        pointRx pPointRx[2] = {x=594.549819, y=30.770866, z=171.45682, rx=-40.410864, ry=94.502866, rz=40.920287, shoulder=lefty, elbow=epositive, wrist=wnegative}
        string sID
      [28]
        bool bMarked
        jointRx jJointRx = {j1=-1.639134, j2=22.193742, j3=116.03978, j4=1.817031, j5=-44.819098, j6=-0.790246}
        pointRx pInter
        paraItem pParaItem
          [0]
            bool bSafePoint
            ifItem iIfItem
              [0]
                bool bANDOR[2]
                num nSigIndex[3]
                num nSigType[3]
                num nValue[3]
            mdesc mMdesc = {accel=25, vel=50, leave=1}
            num nActionIndex = 8
            num nDelay = 1.2
            num nMoveType = 7
            num nPercentage
            num nSigValue = 1
        pointRx pPointRx[2] = {x=594.549757, y=30.770873, z=70.540177, rx=-40.399083, ry=94.503271, rz=40.908669, shoulder=lefty, elbow=epositive, wrist=wnegative}
        string sID
      [29]
        bool bMarked
        jointRx jJointRx = {j1=-1.639045, j2=12.402747, j3=111.595585, j4=2.517874, j5=-30.594648, j6=-1.669011}
        pointRx pInter
        paraItem pParaItem
          [0]
            bool bSafePoint
            ifItem iIfItem
              [0]
                bool bANDOR[2]
                num nSigIndex[3]
                num nSigType[3]
                num nValue[3]
            mdesc mMdesc
            num nActionIndex = 10
            num nDelay = 5
            num nMoveType = 4
            num nPercentage
            num nSigValue
        pointRx pPointRx[2] = {x=594.549819, y=30.770866, z=171.45682, rx=-40.410864, ry=94.502866, rz=40.920287, shoulder=lefty, elbow=epositive, wrist=wnegative}
        string sID
      [30]
        bool bMarked
        jointRx jJointRx = {j1=-1.639045, j2=12.402747, j3=111.595585, j4=2.517874, j5=-30.594648, j6=-1.669011}
        pointRx pInter
        paraItem pParaItem
          [0]
            bool bSafePoint
            ifItem iIfItem
              [0]
                bool bANDOR[2]
                num nSigIndex[3]
                num nSigType[3]
                num nValue[3]
            mdesc mMdesc
            num nActionIndex = 10
            num nDelay = 0.5
            num nMoveType = 7
            num nPercentage
            num nSigValue
        pointRx pPointRx[2] = {x=594.549819, y=30.770866, z=171.45682, rx=-40.410864, ry=94.502866, rz=40.920287, shoulder=lefty, elbow=epositive, wrist=wnegative}
        string sID
      [31]
        bool bMarked
        jointRx jJointRx = {j1=-1.639045, j2=12.402747, j3=111.595585, j4=2.517874, j5=-30.594648, j6=-1.669011}
        pointRx pInter
        paraItem pParaItem
          [0]
            bool bSafePoint
            ifItem iIfItem
              [0]
                bool bANDOR[2]
                num nSigIndex[3]
                num nSigType[3]
                num nValue[3]
            mdesc mMdesc
            num nActionIndex = 9
            num nDelay = 5
            num nMoveType = 3
            num nPercentage
            num nSigValue = 1
        pointRx pPointRx[2] = {x=594.549819, y=30.770866, z=171.45682, rx=-40.410864, ry=94.502866, rz=40.920287, shoulder=lefty, elbow=epositive, wrist=wnegative}
        string sID
      [32]
        bool bMarked
        jointRx jJointRx = {j1=-7.226415, j2=23.592658, j3=117.966616, j4=-6.814076, j5=-74.706283, j6=4.672196}
        pointRx pInter
        paraItem pParaItem
          [0]
            bool bSafePoint
            ifItem iIfItem
              [0]
                bool bANDOR[2]
                num nSigIndex[3]
                num nSigType[3]
                num nValue[3]
            mdesc mMdesc
            num nActionIndex = 9
            num nDelay = 5
            num nMoveType
            num nPercentage
            num nSigValue = 1
        pointRx pPointRx[2] = {x=578.895133, y=-11.466034, z=95.479539, rx=0.214531, ry=67.116514, rz=-0.152975, shoulder=lefty, elbow=epositive, wrist=wnegative}
        string sID
      [33]
        bool bMarked
        jointRx jJointRx = {j1=-2.687248, j2=16.117165, j3=122.304638, j4=-0.487867, j5=-66.528565, j6=1.978834}
        pointRx pInter
        paraItem pParaItem
          [0]
            bool bSafePoint
            ifItem iIfItem
              [0]
                bool bANDOR[2]
                num nSigIndex[3]
                num nSigType[3]
                num nValue[3]
            mdesc mMdesc
            num nActionIndex = 1
            num nDelay = 5
            num nMoveType = 6
            num nPercentage
            num nSigValue = 1
        pointRx pPointRx[2] = {x=546.855577, y=25.169852, z=121.450925, rx=6.745985, ry=71.76392, rz=-5.460967, shoulder=lefty, elbow=epositive, wrist=wnegative}
        string sID
      [34]
        bool bMarked
        jointRx jJointRx = {j1=-2.687248, j2=16.117165, j3=122.304638, j4=-0.487867, j5=-66.528565, j6=1.978834}
        pointRx pInter
        paraItem pParaItem
          [0]
            bool bSafePoint
            ifItem iIfItem
              [0]
                bool bANDOR[2]
                num nSigIndex[3]
                num nSigType[3]
                num nValue[3]
            mdesc mMdesc
            num nActionIndex = 1
            num nDelay = 5
            num nMoveType = 5
            num nPercentage
            num nSigValue = 1
        pointRx pPointRx[2] = {x=546.855577, y=25.169852, z=121.450925, rx=6.745985, ry=71.76392, rz=-5.460967, shoulder=lefty, elbow=epositive, wrist=wnegative}
        string sID
      [35]
        bool bMarked
        jointRx jJointRx = {j1=-1.639045, j2=12.402747, j3=111.595585, j4=2.517874, j5=-30.594648, j6=-1.669011}
        pointRx pInter
        paraItem pParaItem
          [0]
            bool bSafePoint
            ifItem iIfItem
              [0]
                bool bANDOR[2]
                num nSigIndex[3]
                num nSigType[3]
                num nValue[3]
            mdesc mMdesc
            num nActionIndex = 10
            num nDelay
            num nMoveType = 4
            num nPercentage
            num nSigValue = 1
        pointRx pPointRx[2] = {x=594.549819, y=30.770866, z=171.45682, rx=-40.410864, ry=94.502866, rz=40.920287, shoulder=lefty, elbow=epositive, wrist=wnegative}
        string sID
      [36]
        bool bMarked
        jointRx jJointRx = {j1=-1.639045, j2=12.402747, j3=111.595585, j4=2.517874, j5=-30.594648, j6=-1.669011}
        pointRx pInter
        paraItem pParaItem
          [0]
            bool bSafePoint
            ifItem iIfItem
              [0]
                bool bANDOR[2]
                num nSigIndex[3]
                num nSigType[3]
                num nValue[3]
            mdesc mMdesc
            num nActionIndex = 8
            num nDelay
            num nMoveType = 3
            num nPercentage
            num nSigValue = 1
        pointRx pPointRx[2] = {x=594.549819, y=30.770866, z=171.45682, rx=-40.410864, ry=94.502866, rz=40.920287, shoulder=lefty, elbow=epositive, wrist=wnegative}
        string sID
      [37]
        bool bMarked
        jointRx jJointRx = {j1=-1.639134, j2=22.193742, j3=116.03978, j4=1.817031, j5=-44.819098, j6=-0.790246}
        pointRx pInter
        paraItem pParaItem
          [0]
            bool bSafePoint
            ifItem iIfItem
              [0]
                bool bANDOR[2]
                num nSigIndex[3]
                num nSigType[3]
                num nValue[3]
            mdesc mMdesc = {accel=25, vel=50, leave=1}
            num nActionIndex = 8
            num nDelay = 1.2
            num nMoveType = 7
            num nPercentage
            num nSigValue = 1
        pointRx pPointRx[2] = {x=594.549757, y=30.770873, z=70.540177, rx=-40.399083, ry=94.503271, rz=40.908669, shoulder=lefty, elbow=epositive, wrist=wnegative}
        string sID
      [38]
        bool bMarked
        jointRx jJointRx = {j1=-1.639045, j2=12.402747, j3=111.595585, j4=2.517874, j5=-30.594648, j6=-1.669011}
        pointRx pInter
        paraItem pParaItem
          [0]
            bool bSafePoint
            ifItem iIfItem
              [0]
                bool bANDOR[2]
                num nSigIndex[3]
                num nSigType[3]
                num nValue[3]
            mdesc mMdesc
            num nActionIndex = 10
            num nDelay = 5
            num nMoveType = 4
            num nPercentage
            num nSigValue
        pointRx pPointRx[2] = {x=594.549819, y=30.770866, z=171.45682, rx=-40.410864, ry=94.502866, rz=40.920287, shoulder=lefty, elbow=epositive, wrist=wnegative}
        string sID
      [39]
        bool bMarked
        jointRx jJointRx = {j1=-1.639045, j2=12.402747, j3=111.595585, j4=2.517874, j5=-30.594648, j6=-1.669011}
        pointRx pInter
        paraItem pParaItem
          [0]
            bool bSafePoint
            ifItem iIfItem
              [0]
                bool bANDOR[2]
                num nSigIndex[3]
                num nSigType[3]
                num nValue[3]
            mdesc mMdesc
            num nActionIndex = 10
            num nDelay = 0.5
            num nMoveType = 7
            num nPercentage
            num nSigValue
        pointRx pPointRx[2] = {x=594.549819, y=30.770866, z=171.45682, rx=-40.410864, ry=94.502866, rz=40.920287, shoulder=lefty, elbow=epositive, wrist=wnegative}
        string sID
      [40]
        bool bMarked
        jointRx jJointRx = {j1=-1.639045, j2=12.402747, j3=111.595585, j4=2.517874, j5=-30.594648, j6=-1.669011}
        pointRx pInter
        paraItem pParaItem
          [0]
            bool bSafePoint
            ifItem iIfItem
              [0]
                bool bANDOR[2]
                num nSigIndex[3]
                num nSigType[3]
                num nValue[3]
            mdesc mMdesc
            num nActionIndex = 9
            num nDelay = 5
            num nMoveType = 3
            num nPercentage
            num nSigValue = 1
        pointRx pPointRx[2] = {x=594.549819, y=30.770866, z=171.45682, rx=-40.410864, ry=94.502866, rz=40.920287, shoulder=lefty, elbow=epositive, wrist=wnegative}
        string sID
      [41]
        bool bMarked
        jointRx jJointRx = {j1=-5.695731, j2=1.0651158, j3=140.857781, j4=-5.0995594, j5=-70.16665, j6=4.945113}
        pointRx pInter
        paraItem pParaItem
          [0]
            bool bSafePoint
            ifItem iIfItem
              [0]
                bool bANDOR[2]
                num nSigIndex[3]
                num nSigType[3]
                num nValue[3]
            mdesc mMdesc
            num nActionIndex = 9
            num nDelay = 5
            num nMoveType
            num nPercentage
            num nSigValue = 1
        pointRx pPointRx[2] = {x=418.431788, y=16.917425, z=121.450805, rx=1.98388, ry=71.88349, rz=-0.448462, shoulder=lefty, elbow=epositive, wrist=wnegative}
        string sID
      [42]
        bool bMarked
        jointRx jJointRx = {j1=-7.298028, j2=2.858926, j3=83.785178, j4=10.154119, j5=40.0244602, j6=-11.233253}
        pointRx pInter
        paraItem pParaItem
          [0]
            bool bSafePoint
            ifItem iIfItem
              [0]
                bool bANDOR[2]
                num nSigIndex[3]
                num nSigType[3]
                num nValue[3]
            mdesc mMdesc
            num nActionIndex = 9
            num nDelay = 5
            num nMoveType
            num nPercentage
            num nSigValue = 1
        pointRx pPointRx[2] = {x=578.748864, y=-12.280333, z=390.636728, rx=1.0385678, ry=125.960392, rz=0.0408503, shoulder=lefty, elbow=epositive, wrist=wpositive}
        string sID
      [43]
        bool bMarked
        jointRx jJointRx = {j1=-11.714441, j2=6.765338, j3=77.722005, j4=11.0036166, j5=46.0689495, j6=-14.380804}
        pointRx pInter
        paraItem pParaItem
          [0]
            bool bSafePoint
            ifItem iIfItem
              [0]
                bool bANDOR[2]
                num nSigIndex[3]
                num nSigType[3]
                num nValue[3]
            mdesc mMdesc
            num nActionIndex = 1
            num nDelay = 5
            num nMoveType = 6
            num nPercentage
            num nSigValue = 1
        pointRx pPointRx[2] = {x=599.417794, y=-59.189006, z=399.167028, rx=-1.744645, ry=129.591612, rz=2.151169, shoulder=lefty, elbow=epositive, wrist=wpositive}
        string sID
      [44]
        bool bMarked
        jointRx jJointRx = {j1=-11.714441, j2=6.765338, j3=77.722005, j4=11.0036166, j5=46.0689495, j6=-14.380804}
        pointRx pInter
        paraItem pParaItem
          [0]
            bool bSafePoint
            ifItem iIfItem
              [0]
                bool bANDOR[2]
                num nSigIndex[3]
                num nSigType[3]
                num nValue[3]
            mdesc mMdesc
            num nActionIndex = 1
            num nDelay = 5
            num nMoveType = 5
            num nPercentage
            num nSigValue = 1
        pointRx pPointRx[2] = {x=599.417794, y=-59.189006, z=399.167028, rx=-1.744645, ry=129.591612, rz=2.151169, shoulder=lefty, elbow=epositive, wrist=wpositive}
        string sID
      [45]
        bool bMarked
        jointRx jJointRx = {j1=-11.714441, j2=6.765338, j3=77.722005, j4=11.0036166, j5=46.0689495, j6=-14.380804}
        pointRx pInter
        paraItem pParaItem
          [0]
            bool bSafePoint
            ifItem iIfItem
              [0]
                bool bANDOR[2]
                num nSigIndex[3]
                num nSigType[3]
                num nValue[3]
            mdesc mMdesc
            num nActionIndex = 10
            num nDelay = 5
            num nMoveType = 4
            num nPercentage
            num nSigValue = 1
        pointRx pPointRx[2] = {x=599.417794, y=-59.189006, z=399.167028, rx=-1.744645, ry=129.591612, rz=2.151169, shoulder=lefty, elbow=epositive, wrist=wpositive}
        string sID
      [46]
        bool bMarked
        jointRx jJointRx = {j1=-11.714441, j2=6.765338, j3=77.722005, j4=11.0036166, j5=46.0689495, j6=-14.380804}
        pointRx pInter
        paraItem pParaItem
          [0]
            bool bSafePoint
            ifItem iIfItem
              [0]
                bool bANDOR[2]
                num nSigIndex[3]
                num nSigType[3]
                num nValue[3]
            mdesc mMdesc
            num nActionIndex = 8
            num nDelay = 5
            num nMoveType = 3
            num nPercentage
            num nSigValue = 1
        pointRx pPointRx[2] = {x=599.417794, y=-59.189006, z=399.167028, rx=-1.744645, ry=129.591612, rz=2.151169, shoulder=lefty, elbow=epositive, wrist=wpositive}
        string sID
      [47]
        bool bMarked
        jointRx jJointRx = {j1=-11.714441, j2=6.765338, j3=77.722005, j4=11.0036166, j5=46.0689495, j6=-14.380804}
        pointRx pInter
        paraItem pParaItem
          [0]
            bool bSafePoint
            ifItem iIfItem
              [0]
                bool bANDOR[2]
                num nSigIndex[3]
                num nSigType[3]
                num nValue[3]
            mdesc mMdesc
            num nActionIndex = 8
            num nDelay = 2
            num nMoveType = 7
            num nPercentage
            num nSigValue = 1
        pointRx pPointRx[2] = {x=599.417794, y=-59.189006, z=399.167028, rx=-1.744645, ry=129.591612, rz=2.151169, shoulder=lefty, elbow=epositive, wrist=wpositive}
        string sID
      [48]
        bool bMarked
        jointRx jJointRx = {j1=-11.714441, j2=6.765338, j3=77.722005, j4=11.0036166, j5=46.0689495, j6=-14.380804}
        pointRx pInter
        paraItem pParaItem
          [0]
            bool bSafePoint
            ifItem iIfItem
              [0]
                bool bANDOR[2]
                num nSigIndex[3]
                num nSigType[3]
                num nValue[3]
            mdesc mMdesc
            num nActionIndex = 10
            num nDelay = 1
            num nMoveType = 4
            num nPercentage
            num nSigValue
        pointRx pPointRx[2] = {x=599.417794, y=-59.189006, z=399.167028, rx=-1.744645, ry=129.591612, rz=2.151169, shoulder=lefty, elbow=epositive, wrist=wpositive}
        string sID
      [49]
        bool bMarked
        jointRx jJointRx = {j1=-11.714441, j2=6.765338, j3=77.722005, j4=11.0036166, j5=46.0689495, j6=-14.380804}
        pointRx pInter
        paraItem pParaItem
          [0]
            bool bSafePoint
            ifItem iIfItem
              [0]
                bool bANDOR[2]
                num nSigIndex[3]
                num nSigType[3]
                num nValue[3]
            mdesc mMdesc
            num nActionIndex = 10
            num nDelay = 0.5
            num nMoveType = 7
            num nPercentage
            num nSigValue
        pointRx pPointRx[2] = {x=599.417794, y=-59.189006, z=399.167028, rx=-1.744645, ry=129.591612, rz=2.151169, shoulder=lefty, elbow=epositive, wrist=wpositive}
        string sID
      [50]
        bool bMarked
        jointRx jJointRx = {j1=-11.714441, j2=6.765338, j3=77.722005, j4=11.0036166, j5=46.0689495, j6=-14.380804}
        pointRx pInter
        paraItem pParaItem
          [0]
            bool bSafePoint
            ifItem iIfItem
              [0]
                bool bANDOR[2]
                num nSigIndex[3]
                num nSigType[3]
                num nValue[3]
            mdesc mMdesc
            num nActionIndex = 9
            num nDelay = 1
            num nMoveType = 3
            num nPercentage
            num nSigValue = 1
        pointRx pPointRx[2] = {x=599.417794, y=-59.189006, z=399.167028, rx=-1.744645, ry=129.591612, rz=2.151169, shoulder=lefty, elbow=epositive, wrist=wpositive}
        string sID
      [51]
        bool bMarked
        jointRx jJointRx = {j1=-1.121423, j2=3.0557806, j3=83.578223, j4=2.394681, j5=39.358319, j6=-1.629384}
        pointRx pInter
        paraItem pParaItem
          [0]
            bool bSafePoint
            ifItem iIfItem
              [0]
                bool bANDOR[2]
                num nSigIndex[3]
                num nSigType[3]
                num nValue[3]
            mdesc mMdesc
            num nActionIndex = 9
            num nDelay = 5
            num nMoveType
            num nPercentage
            num nSigValue = 1
        pointRx pPointRx[2] = {x=578.748846, y=41.330803, z=390.636723, rx=1.0399619, ry=125.960028, rz=0.0394555, shoulder=lefty, elbow=epositive, wrist=wpositive}
        string sID
      [52]
        bool bMarked
        jointRx jJointRx = {j1=-2.687248, j2=16.117165, j3=122.304638, j4=-0.487867, j5=-66.528565, j6=1.978834}
        pointRx pInter
        paraItem pParaItem
          [0]
            bool bSafePoint
            ifItem iIfItem
              [0]
                bool bANDOR[2]
                num nSigIndex[3]
                num nSigType[3]
                num nValue[3]
            mdesc mMdesc
            num nActionIndex = 1
            num nDelay = 5
            num nMoveType = 6
            num nPercentage
            num nSigValue = 1
        pointRx pPointRx[2] = {x=546.855577, y=25.169852, z=121.450925, rx=6.745985, ry=71.76392, rz=-5.460967, shoulder=lefty, elbow=epositive, wrist=wnegative}
        string sID
      [53]
        bool bMarked
        jointRx jJointRx = {j1=-2.687248, j2=16.117165, j3=122.304638, j4=-0.487867, j5=-66.528565, j6=1.978834}
        pointRx pInter
        paraItem pParaItem
          [0]
            bool bSafePoint
            ifItem iIfItem
              [0]
                bool bANDOR[2]
                num nSigIndex[3]
                num nSigType[3]
                num nValue[3]
            mdesc mMdesc
            num nActionIndex = 1
            num nDelay = 5
            num nMoveType = 5
            num nPercentage
            num nSigValue = 1
        pointRx pPointRx[2] = {x=546.855577, y=25.169852, z=121.450925, rx=6.745985, ry=71.76392, rz=-5.460967, shoulder=lefty, elbow=epositive, wrist=wnegative}
        string sID
      [54]
        bool bMarked
        jointRx jJointRx = {j1=-1.639045, j2=12.402747, j3=111.595585, j4=2.517874, j5=-30.594648, j6=-1.669011}
        pointRx pInter
        paraItem pParaItem
          [0]
            bool bSafePoint
            ifItem iIfItem
              [0]
                bool bANDOR[2]
                num nSigIndex[3]
                num nSigType[3]
                num nValue[3]
            mdesc mMdesc
            num nActionIndex = 10
            num nDelay
            num nMoveType = 4
            num nPercentage
            num nSigValue = 1
        pointRx pPointRx[2] = {x=594.549819, y=30.770866, z=171.45682, rx=-40.410864, ry=94.502866, rz=40.920287, shoulder=lefty, elbow=epositive, wrist=wnegative}
        string sID
      [55]
        bool bMarked
        jointRx jJointRx = {j1=-1.639045, j2=12.402747, j3=111.595585, j4=2.517874, j5=-30.594648, j6=-1.669011}
        pointRx pInter
        paraItem pParaItem
          [0]
            bool bSafePoint
            ifItem iIfItem
              [0]
                bool bANDOR[2]
                num nSigIndex[3]
                num nSigType[3]
                num nValue[3]
            mdesc mMdesc
            num nActionIndex = 8
            num nDelay
            num nMoveType = 3
            num nPercentage
            num nSigValue = 1
        pointRx pPointRx[2] = {x=594.549819, y=30.770866, z=171.45682, rx=-40.410864, ry=94.502866, rz=40.920287, shoulder=lefty, elbow=epositive, wrist=wnegative}
        string sID
      [56]
        bool bMarked
        jointRx jJointRx = {j1=-1.639134, j2=22.193742, j3=116.03978, j4=1.817031, j5=-44.819098, j6=-0.790246}
        pointRx pInter
        paraItem pParaItem
          [0]
            bool bSafePoint
            ifItem iIfItem
              [0]
                bool bANDOR[2]
                num nSigIndex[3]
                num nSigType[3]
                num nValue[3]
            mdesc mMdesc = {accel=25, vel=50, leave=1}
            num nActionIndex = 8
            num nDelay = 2
            num nMoveType = 7
            num nPercentage
            num nSigValue = 1
        pointRx pPointRx[2] = {x=594.549757, y=30.770873, z=70.540177, rx=-40.399083, ry=94.503271, rz=40.908669, shoulder=lefty, elbow=epositive, wrist=wnegative}
        string sID
      [57]
        bool bMarked
        jointRx jJointRx = {j1=-1.639045, j2=12.402747, j3=111.595585, j4=2.517874, j5=-30.594648, j6=-1.669011}
        pointRx pInter
        paraItem pParaItem
          [0]
            bool bSafePoint
            ifItem iIfItem
              [0]
                bool bANDOR[2]
                num nSigIndex[3]
                num nSigType[3]
                num nValue[3]
            mdesc mMdesc
            num nActionIndex = 10
            num nDelay = 5
            num nMoveType = 4
            num nPercentage
            num nSigValue
        pointRx pPointRx[2] = {x=594.549819, y=30.770866, z=171.45682, rx=-40.410864, ry=94.502866, rz=40.920287, shoulder=lefty, elbow=epositive, wrist=wnegative}
        string sID
      [58]
        bool bMarked
        jointRx jJointRx = {j1=-1.639045, j2=12.402747, j3=111.595585, j4=2.517874, j5=-30.594648, j6=-1.669011}
        pointRx pInter
        paraItem pParaItem
          [0]
            bool bSafePoint
            ifItem iIfItem
              [0]
                bool bANDOR[2]
                num nSigIndex[3]
                num nSigType[3]
                num nValue[3]
            mdesc mMdesc
            num nActionIndex = 10
            num nDelay = 0.5
            num nMoveType = 7
            num nPercentage
            num nSigValue
        pointRx pPointRx[2] = {x=594.549819, y=30.770866, z=171.45682, rx=-40.410864, ry=94.502866, rz=40.920287, shoulder=lefty, elbow=epositive, wrist=wnegative}
        string sID
      [59]
        bool bMarked
        jointRx jJointRx = {j1=-1.639045, j2=12.402747, j3=111.595585, j4=2.517874, j5=-30.594648, j6=-1.669011}
        pointRx pInter
        paraItem pParaItem
          [0]
            bool bSafePoint
            ifItem iIfItem
              [0]
                bool bANDOR[2]
                num nSigIndex[3]
                num nSigType[3]
                num nValue[3]
            mdesc mMdesc
            num nActionIndex = 9
            num nDelay = 5
            num nMoveType = 3
            num nPercentage
            num nSigValue = 1
        pointRx pPointRx[2] = {x=594.549819, y=30.770866, z=171.45682, rx=-40.410864, ry=94.502866, rz=40.920287, shoulder=lefty, elbow=epositive, wrist=wnegative}
        string sID
      [60]
        bool bMarked
        jointRx jJointRx = {j1=-3.420163, j2=22.945404, j3=44.641192, j4=2.309583, j5=82.959552, j6=-2.373603}
        pointRx pInter
        paraItem pParaItem
          [0]
            bool bSafePoint
            ifItem iIfItem
              [0]
                bool bANDOR[2]
                num nSigIndex[3]
                num nSigType[3]
                num nValue[3]
            mdesc mMdesc
            num nActionIndex = 9
            num nDelay = 5
            num nMoveType
            num nPercentage
            num nSigValue = 1
        pointRx pPointRx[2] = {x=659.773544, y=14.665083, z=466.418783, rx=0.698518, ry=150.466936, rz=0.542991, shoulder=lefty, elbow=epositive, wrist=wpositive}
        string sID
      [61]
        bool bMarked
        jointRx jJointRx = {j1=-2.687248, j2=16.117165, j3=122.304638, j4=-0.487867, j5=-66.528565, j6=1.978834}
        pointRx pInter
        paraItem pParaItem
          [0]
            bool bSafePoint
            ifItem iIfItem
              [0]
                bool bANDOR[2]
                num nSigIndex[3]
                num nSigType[3]
                num nValue[3]
            mdesc mMdesc
            num nActionIndex = 1
            num nDelay = 5
            num nMoveType = 6
            num nPercentage
            num nSigValue = 1
        pointRx pPointRx[2] = {x=546.855577, y=25.169852, z=121.450925, rx=6.745985, ry=71.76392, rz=-5.460967, shoulder=lefty, elbow=epositive, wrist=wnegative}
        string sID
      [62]
        bool bMarked
        jointRx jJointRx = {j1=-2.687248, j2=16.117165, j3=122.304638, j4=-0.487867, j5=-66.528565, j6=1.978834}
        pointRx pInter
        paraItem pParaItem
          [0]
            bool bSafePoint
            ifItem iIfItem
              [0]
                bool bANDOR[2]
                num nSigIndex[3]
                num nSigType[3]
                num nValue[3]
            mdesc mMdesc
            num nActionIndex = 1
            num nDelay = 5
            num nMoveType = 5
            num nPercentage
            num nSigValue = 1
        pointRx pPointRx[2] = {x=546.855577, y=25.169852, z=121.450925, rx=6.745985, ry=71.76392, rz=-5.460967, shoulder=lefty, elbow=epositive, wrist=wnegative}
        string sID
      [63]
        bool bMarked
        jointRx jJointRx = {j1=-1.639045, j2=12.402747, j3=111.595585, j4=2.517874, j5=-30.594648, j6=-1.669011}
        pointRx pInter
        paraItem pParaItem
          [0]
            bool bSafePoint
            ifItem iIfItem
              [0]
                bool bANDOR[2]
                num nSigIndex[3]
                num nSigType[3]
                num nValue[3]
            mdesc mMdesc
            num nActionIndex = 10
            num nDelay
            num nMoveType = 4
            num nPercentage
            num nSigValue = 1
        pointRx pPointRx[2] = {x=594.549819, y=30.770866, z=171.45682, rx=-40.410864, ry=94.502866, rz=40.920287, shoulder=lefty, elbow=epositive, wrist=wnegative}
        string sID
      [64]
        bool bMarked
        jointRx jJointRx = {j1=-1.639045, j2=12.402747, j3=111.595585, j4=2.517874, j5=-30.594648, j6=-1.669011}
        pointRx pInter
        paraItem pParaItem
          [0]
            bool bSafePoint
            ifItem iIfItem
              [0]
                bool bANDOR[2]
                num nSigIndex[3]
                num nSigType[3]
                num nValue[3]
            mdesc mMdesc
            num nActionIndex = 8
            num nDelay
            num nMoveType = 3
            num nPercentage
            num nSigValue = 1
        pointRx pPointRx[2] = {x=594.549819, y=30.770866, z=171.45682, rx=-40.410864, ry=94.502866, rz=40.920287, shoulder=lefty, elbow=epositive, wrist=wnegative}
        string sID
      [65]
        bool bMarked
        jointRx jJointRx = {j1=-1.639134, j2=22.193742, j3=116.03978, j4=1.817031, j5=-44.819098, j6=-0.790246}
        pointRx pInter
        paraItem pParaItem
          [0]
            bool bSafePoint
            ifItem iIfItem
              [0]
                bool bANDOR[2]
                num nSigIndex[3]
                num nSigType[3]
                num nValue[3]
            mdesc mMdesc = {accel=25, vel=50, leave=1}
            num nActionIndex = 8
            num nDelay = 1.2
            num nMoveType = 7
            num nPercentage
            num nSigValue = 1
        pointRx pPointRx[2] = {x=594.549757, y=30.770873, z=70.540177, rx=-40.399083, ry=94.503271, rz=40.908669, shoulder=lefty, elbow=epositive, wrist=wnegative}
        string sID
      [66]
        bool bMarked
        jointRx jJointRx = {j1=-1.639045, j2=12.402747, j3=111.595585, j4=2.517874, j5=-30.594648, j6=-1.669011}
        pointRx pInter
        paraItem pParaItem
          [0]
            bool bSafePoint
            ifItem iIfItem
              [0]
                bool bANDOR[2]
                num nSigIndex[3]
                num nSigType[3]
                num nValue[3]
            mdesc mMdesc
            num nActionIndex = 10
            num nDelay = 5
            num nMoveType = 4
            num nPercentage
            num nSigValue
        pointRx pPointRx[2] = {x=594.549819, y=30.770866, z=171.45682, rx=-40.410864, ry=94.502866, rz=40.920287, shoulder=lefty, elbow=epositive, wrist=wnegative}
        string sID
      [67]
        bool bMarked
        jointRx jJointRx = {j1=-1.639045, j2=12.402747, j3=111.595585, j4=2.517874, j5=-30.594648, j6=-1.669011}
        pointRx pInter
        paraItem pParaItem
          [0]
            bool bSafePoint
            ifItem iIfItem
              [0]
                bool bANDOR[2]
                num nSigIndex[3]
                num nSigType[3]
                num nValue[3]
            mdesc mMdesc
            num nActionIndex = 10
            num nDelay = 0.5
            num nMoveType = 7
            num nPercentage
            num nSigValue
        pointRx pPointRx[2] = {x=594.549819, y=30.770866, z=171.45682, rx=-40.410864, ry=94.502866, rz=40.920287, shoulder=lefty, elbow=epositive, wrist=wnegative}
        string sID
      [68]
        bool bMarked
        jointRx jJointRx = {j1=-1.639045, j2=12.402747, j3=111.595585, j4=2.517874, j5=-30.594648, j6=-1.669011}
        pointRx pInter
        paraItem pParaItem
          [0]
            bool bSafePoint
            ifItem iIfItem
              [0]
                bool bANDOR[2]
                num nSigIndex[3]
                num nSigType[3]
                num nValue[3]
            mdesc mMdesc
            num nActionIndex = 9
            num nDelay = 5
            num nMoveType = 3
            num nPercentage
            num nSigValue = 1
        pointRx pPointRx[2] = {x=594.549819, y=30.770866, z=171.45682, rx=-40.410864, ry=94.502866, rz=40.920287, shoulder=lefty, elbow=epositive, wrist=wnegative}
        string sID
      [69]
        bool bMarked
        jointRx jJointRx = {j1=-5.00727366, j2=-18.178881, j3=100.185408, j4=3.718834, j5=47.673508, j6=-4.893046}
        pointRx pInter
        paraItem pParaItem
          [0]
            bool bSafePoint
            ifItem iIfItem
              [0]
                bool bANDOR[2]
                num nSigIndex[3]
                num nSigType[3]
                num nValue[3]
            mdesc mMdesc
            num nActionIndex = 9
            num nDelay = 5
            num nMoveType
            num nPercentage
            num nSigValue = 1
        pointRx pPointRx[2] = {x=418.415736, y=18.345016, z=399.191838, rx=-1.743265, ry=129.587286, rz=2.147877, shoulder=lefty, elbow=epositive, wrist=wpositive}
        string sID
      [70]
        bool bMarked
        jointRx jJointRx = {j1=-1.296156, j2=5.897159, j3=133.210861, j4=1.250253, j5=-71.161646, j6=1.72109}
        pointRx pInter
        paraItem pParaItem
          [0]
            bool bSafePoint
            ifItem iIfItem
              [0]
                bool bANDOR[2]
                num nSigIndex[3]
                num nSigType[3]
                num nValue[3]
            mdesc mMdesc
            num nActionIndex = 9
            num nDelay = 5
            num nMoveType
            num nPercentage
            num nSigValue = 1
        pointRx pPointRx[2] = {x=465.517432, y=37.4144, z=139.00686202, rx=6.325655, ry=67.813303, rz=-4.2228, shoulder=lefty, elbow=epositive, wrist=wnegative}
        string sID
      [71]
        bool bMarked
        jointRx jJointRx = {j1=-11.359718, j2=15.689869, j3=118.29756, j4=-11.285106, j5=-66.838302, j6=10.0776989}
        pointRx pInter
        paraItem pParaItem
          [0]
            bool bSafePoint
            ifItem iIfItem
              [0]
                bool bANDOR[2]
                num nSigIndex[3]
                num nSigType[3]
                num nValue[3]
            mdesc mMdesc
            num nActionIndex = 9
            num nDelay = 5
            num nMoveType
            num nPercentage
            num nSigValue = 1
        pointRx pPointRx[2] = {x=564.0240975, y=-43.964202, z=151.556021, rx=0.409564, ry=67.941454, rz=0.897692, shoulder=lefty, elbow=epositive, wrist=wnegative}
        string sID
      [72]
        bool bMarked
        jointRx jJointRx = {j1=-2.687248, j2=16.117165, j3=122.304638, j4=-0.487867, j5=-66.528565, j6=1.978834}
        pointRx pInter
        paraItem pParaItem
          [0]
            bool bSafePoint
            ifItem iIfItem
              [0]
                bool bANDOR[2]
                num nSigIndex[3]
                num nSigType[3]
                num nValue[3]
            mdesc mMdesc
            num nActionIndex = 1
            num nDelay = 5
            num nMoveType = 6
            num nPercentage
            num nSigValue = 1
        pointRx pPointRx[2] = {x=546.855577, y=25.169852, z=121.450925, rx=6.745985, ry=71.76392, rz=-5.460967, shoulder=lefty, elbow=epositive, wrist=wnegative}
        string sID
      [73]
        bool bMarked
        jointRx jJointRx = {j1=-2.687248, j2=16.117165, j3=122.304638, j4=-0.487867, j5=-66.528565, j6=1.978834}
        pointRx pInter
        paraItem pParaItem
          [0]
            bool bSafePoint
            ifItem iIfItem
              [0]
                bool bANDOR[2]
                num nSigIndex[3]
                num nSigType[3]
                num nValue[3]
            mdesc mMdesc
            num nActionIndex = 1
            num nDelay = 5
            num nMoveType = 5
            num nPercentage
            num nSigValue = 1
        pointRx pPointRx[2] = {x=546.855577, y=25.169852, z=121.450925, rx=6.745985, ry=71.76392, rz=-5.460967, shoulder=lefty, elbow=epositive, wrist=wnegative}
        string sID
      [74]
        bool bMarked
        jointRx jJointRx = {j1=-1.639045, j2=12.402747, j3=111.595585, j4=2.517874, j5=-30.594648, j6=-1.669011}
        pointRx pInter
        paraItem pParaItem
          [0]
            bool bSafePoint
            ifItem iIfItem
              [0]
                bool bANDOR[2]
                num nSigIndex[3]
                num nSigType[3]
                num nValue[3]
            mdesc mMdesc
            num nActionIndex = 10
            num nDelay
            num nMoveType = 4
            num nPercentage
            num nSigValue = 1
        pointRx pPointRx[2] = {x=594.549819, y=30.770866, z=171.45682, rx=-40.410864, ry=94.502866, rz=40.920287, shoulder=lefty, elbow=epositive, wrist=wnegative}
        string sID
      [75]
        bool bMarked
        jointRx jJointRx = {j1=-1.639045, j2=12.402747, j3=111.595585, j4=2.517874, j5=-30.594648, j6=-1.669011}
        pointRx pInter
        paraItem pParaItem
          [0]
            bool bSafePoint
            ifItem iIfItem
              [0]
                bool bANDOR[2]
                num nSigIndex[3]
                num nSigType[3]
